(* IEC 61131-3 sources: helmsman/crates/helmsman-node/bench, 7 files *)

(* ---- analog_scale.st ---- *)
(* Raw analog count to engineering units, held to the range. bad is set when
   the raw value is outside raw_min..raw_max by more than the margin: a broken
   wire on a 4-20 mA loop, or a transmitter that has failed. *)
FUNCTION_BLOCK analog_scale
VAR_INPUT
  raw : REAL;
  raw_min : REAL := 0.0;
  raw_max : REAL := 32767.0;
  eng_min : REAL := 0.0;
  eng_max : REAL := 100.0;
  margin : REAL := 0.05;
END_VAR
VAR_OUTPUT
  value : REAL;
  bad : BOOL;
END_VAR
VAR
  span : REAL;
END_VAR
span := raw_max - raw_min;
bad := span <= 0.0 OR raw < raw_min - span * margin OR raw > raw_max + span * margin;
IF span > 0.0 THEN
  value := LIMIT(eng_min, eng_min + (raw - raw_min) / span * (eng_max - eng_min), eng_max);
END_IF;
END_FUNCTION_BLOCK

(* ---- batch_mixer.st ---- *)
(* Batch mixing tank: fill, heat while agitating, hold, drain, repeat.

   plant_model.st stands in for the tank so this runs with nothing wired. To
   wire real I/O: delete plant_model.st, delete the plant lines in the PROGRAM
   (each one says PLANT), and point io.map at your remote I/O module.

   A heater and agitator need a hardwired over-temperature cut-out and E-stop
   circuit. Those belong in hardware; nothing here is a safety function. *)

FUNCTION_BLOCK mixer_tank
VAR_INPUT
  run : BOOL;
  ack : BOOL;
  level_m : REAL;
  temp_c : REAL;
  inlet_open_sw : BOOL;
  inlet_closed_sw : BOOL;
  outlet_open_sw : BOOL;
  outlet_closed_sw : BOOL;
  agitator_fb : BOOL;
  agitator_overload : BOOL;
  overtemp_sw : BOOL;
END_VAR
VAR_OUTPUT
  inlet_coil : BOOL;
  outlet_coil : BOOL;
  agitator_contactor : BOOL;
  heater : BOOL;
  step : INT;
  batches : INT;
  tripped : BOOL;
  alarm_new : BOOL;
END_VAR
VAR CONSTANT
  fill_to_m : REAL := 2.0;        (* batch level *)
  empty_at_m : REAL := 0.05;      (* drained *)
  heater_min_m : REAL := 0.5;     (* element covered *)
  heat_to_c : REAL := 60.0;       (* batch temperature *)
  over_c : REAL := 80.0;          (* high temperature alarm *)
  hold_time : TIME := T#10s;      (* mix at temperature *)
  fill_max : TIME := T#60s;
  heat_max : TIME := T#120s;
  drain_max : TIME := T#60s;
END_VAR
VAR
  seq : step_sequencer;
  inlet : solenoid_valve;
  outlet : solenoid_valve;
  agitator : motor_starter;
  high_temp : latched_alarm;
  step_late : latched_alarm;
  equipment : latched_alarm;
  hold : TON;
  step_done : BOOL;
  step_max : TIME;
  want_inlet : BOOL;
  want_outlet : BOOL;
  want_agitator : BOOL;
  want_heat : BOOL;
END_VAR

high_temp(condition := overtemp_sw OR temp_c >= over_c, ack := ack, on_delay := T#0s);
step_late(condition := seq.timed_out, ack := ack, on_delay := T#0s);
equipment(condition := inlet.fault OR outlet.fault OR agitator.fault, ack := ack, on_delay := T#0s);
tripped := high_temp.showing OR step_late.showing OR equipment.showing;
alarm_new := high_temp.unacked OR step_late.unacked OR equipment.unacked;

seq(start := run AND NOT tripped, advance := step_done, abort := NOT run OR tripped,
    last_step := 4, step_limit := step_max);
step := seq.step;

want_inlet := FALSE;
want_outlet := FALSE;
want_agitator := FALSE;
want_heat := FALSE;
step_done := FALSE;
step_max := T#0s;
CASE step OF
  1: (* fill *)
    want_inlet := level_m < fill_to_m;
    step_done := level_m >= fill_to_m AND inlet.is_closed;
    step_max := fill_max;
  2: (* heat, agitating *)
    want_agitator := TRUE;
    want_heat := agitator.running;
    step_done := temp_c >= heat_to_c;
    step_max := heat_max;
  3: (* hold at temperature *)
    want_agitator := TRUE;
    want_heat := agitator.running AND temp_c < heat_to_c;
    step_done := hold.Q;
  4: (* drain *)
    want_outlet := level_m > empty_at_m;
    step_done := level_m <= empty_at_m AND outlet.is_closed;
    step_max := drain_max;
END_CASE;
hold(IN := step = 3, PT := hold_time);
IF seq.done AND batches < 32767 THEN
  batches := batches + 1;
END_IF;

inlet(open := want_inlet, at_open := inlet_open_sw, at_closed := inlet_closed_sw, reset := ack);
outlet(open := want_outlet, at_open := outlet_open_sw, at_closed := outlet_closed_sw, reset := ack);
agitator(run := want_agitator, feedback := agitator_fb, overload := agitator_overload, reset := ack);
inlet_coil := inlet.coil;
outlet_coil := outlet.coil;
agitator_contactor := agitator.contactor;
(* The heater never runs uncovered, without the agitator, or on an alarm. *)
heater := want_heat AND level_m >= heater_min_m AND NOT tripped;
END_FUNCTION_BLOCK

PROGRAM mixer
VAR_INPUT
  start_pb : BOOL;
  stop_pb : BOOL;
  ack_pb : BOOL;
  inlet_open_in : BOOL;
  inlet_closed_in : BOOL;
  outlet_open_in : BOOL;
  outlet_closed_in : BOOL;
  agitator_fb_in : BOOL;
  agitator_overload_in : BOOL;
  overtemp_in : BOOL;
  sim_inlet_stuck : BOOL;  (* PLANT: the inlet valve never opens *)
END_VAR
VAR_OUTPUT
  inlet_valve : BOOL;
  outlet_valve : BOOL;
  agitator : BOOL;
  heater : BOOL;
  lamp_green : BOOL;
  lamp_red : BOOL;
  step : INT;
  batches : INT;
  level_m : REAL;
  temp_c : REAL;
END_VAR
VAR
  plant : plant_model;  (* PLANT *)
  level_tx : analog_scale;
  temp_tx : analog_scale;
  tank : mixer_tank;
  light : stack_light;
  run : BOOL;
  level_raw : REAL;
  temp_raw : REAL;
  inlet_open : BOOL;
  inlet_closed : BOOL;
  outlet_open : BOOL;
  outlet_closed : BOOL;
  agitator_fb : BOOL;
END_VAR

plant(inlet := inlet_valve, outlet := outlet_valve, agitator := agitator, heater := heater,
      inlet_stuck := sim_inlet_stuck);  (* PLANT *)
level_raw := plant.level_raw;  (* PLANT: read your analog input here *)
temp_raw := plant.temp_raw;    (* PLANT: read your analog input here *)
inlet_open := inlet_open_in OR plant.inlet_open;  (* PLANT: keep the _in input *)
inlet_closed := inlet_closed_in OR plant.inlet_closed;  (* PLANT: keep the _in input *)
outlet_open := outlet_open_in OR plant.outlet_open;  (* PLANT: keep the _in input *)
outlet_closed := outlet_closed_in OR plant.outlet_closed;  (* PLANT: keep the _in input *)
agitator_fb := agitator_fb_in OR plant.agitator_fb;  (* PLANT: keep the _in input *)
run := (run OR start_pb) AND NOT stop_pb AND NOT tank.tripped;

level_tx(raw := level_raw, eng_min := 0.0, eng_max := 3.0);
temp_tx(raw := temp_raw, eng_min := 0.0, eng_max := 120.0);
tank(run := run, ack := ack_pb, level_m := level_tx.value, temp_c := temp_tx.value,
     inlet_open_sw := inlet_open, inlet_closed_sw := inlet_closed,
     outlet_open_sw := outlet_open, outlet_closed_sw := outlet_closed,
     agitator_fb := agitator_fb, agitator_overload := agitator_overload_in,
     overtemp_sw := overtemp_in);
light(running := run, alarm_new := tank.alarm_new, alarm_showing := tank.tripped);

inlet_valve := tank.inlet_coil;
outlet_valve := tank.outlet_coil;
agitator := tank.agitator_contactor;
heater := tank.heater;
lamp_green := light.green;
lamp_red := light.red;
step := tank.step;
batches := tank.batches;
level_m := level_tx.value;
temp_c := temp_tx.value;
END_PROGRAM

(* ---- latched_alarm.st ---- *)
(* One alarm: on after on_delay, stays showing until the condition has gone
   and someone has acknowledged it. *)
FUNCTION_BLOCK latched_alarm
VAR_INPUT
  condition : BOOL;
  ack : BOOL;
  on_delay : TIME;
END_VAR
VAR_OUTPUT
  active : BOOL;
  unacked : BOOL;
  showing : BOOL;
END_VAR
VAR
  delay : TON;
  rise : R_TRIG;
END_VAR
delay(IN := condition, PT := on_delay);
active := delay.Q;
rise(CLK := active);
IF rise.Q THEN
  unacked := TRUE;
ELSIF ack THEN
  unacked := FALSE;
END_IF;
showing := active OR unacked;
END_FUNCTION_BLOCK

(* ---- motor_starter.st ---- *)
(* Motor starter with contactor feedback and a latched fault.
   feedback is the contactor's auxiliary contact, overload the thermal relay.
   fault_code: 0 none, 1 overload, 2 no feedback after a start or feedback
   lost while running, 3 feedback with no command (contactor stuck on).
   A fault drops the contactor and holds until reset. An emergency stop
   belongs in a hardwired safety circuit, not in this block. *)
FUNCTION_BLOCK motor_starter
VAR_INPUT
  run : BOOL;
  feedback : BOOL;
  overload : BOOL;
  reset : BOOL;
  feedback_time : TIME := T#2s;
END_VAR
VAR_OUTPUT
  contactor : BOOL;
  running : BOOL;
  fault : BOOL;
  fault_code : INT;
END_VAR
VAR
  no_feedback : TON;
  stuck_on : TON;
END_VAR
no_feedback(IN := contactor AND NOT feedback, PT := feedback_time);
stuck_on(IN := NOT contactor AND feedback, PT := feedback_time);
IF overload THEN
  fault_code := 1;
ELSIF no_feedback.Q THEN
  fault_code := 2;
ELSIF stuck_on.Q THEN
  fault_code := 3;
ELSIF reset THEN
  fault_code := 0;
END_IF;
fault := fault_code <> 0;
contactor := run AND NOT fault;
running := contactor AND feedback;
END_FUNCTION_BLOCK

(* ---- solenoid_valve.st ---- *)
(* Single-solenoid valve or cylinder with an end switch each way.
   coil follows the command. fault latches when the switch for the commanded
   position has not made within travel_time, and clears on reset once the
   valve has arrived. Both switches on at once counts as not arrived. *)
FUNCTION_BLOCK solenoid_valve
VAR_INPUT
  open : BOOL;
  at_open : BOOL;
  at_closed : BOOL;
  reset : BOOL;
  travel_time : TIME := T#3s;
END_VAR
VAR_OUTPUT
  coil : BOOL;
  is_open : BOOL;
  is_closed : BOOL;
  fault : BOOL;
END_VAR
VAR
  late : TON;
END_VAR
coil := open;
is_open := at_open AND NOT at_closed;
is_closed := at_closed AND NOT at_open;
late(IN := (open AND NOT is_open) OR (NOT open AND NOT is_closed), PT := travel_time);
IF late.Q THEN
  fault := TRUE;
ELSIF reset THEN
  fault := FALSE;
END_IF;
END_FUNCTION_BLOCK

(* ---- stack_light.st ---- *)
(* Green while running. Red flashes for an alarm nobody has acknowledged and
   is steady for one that is acknowledged but still there. *)
FUNCTION_BLOCK stack_light
VAR_INPUT
  running : BOOL;
  alarm_new : BOOL;
  alarm_showing : BOOL;
END_VAR
VAR_OUTPUT
  green : BOOL;
  red : BOOL;
END_VAR
VAR
  flash : BLINK_PATTERN;
  pattern : INT;
END_VAR
IF alarm_new THEN
  pattern := 2;
ELSIF alarm_showing THEN
  pattern := 1;
ELSE
  pattern := 0;
END_IF;
flash(EN := TRUE, MODE := pattern, PERIOD := T#1s);
green := running;
red := flash.Q;
END_FUNCTION_BLOCK

(* ---- step_sequencer.st ---- *)
(* A numbered sequence. Step 0 is idle; start moves to step 1. Each step sets
   advance when it is finished, and the last step goes back to idle with done
   TRUE for one scan. step_limit is how long the current step may take (T#0s:
   no limit); past it, timed_out is set and the step holds until abort. abort
   returns to idle at once. Write the steps in a CASE on the step output. *)
FUNCTION_BLOCK step_sequencer
VAR_INPUT
  start : BOOL;
  advance : BOOL;
  abort : BOOL;
  last_step : INT;
  step_limit : TIME;
END_VAR
VAR_OUTPUT
  step : INT;
  step_time : TIME;
  timed_out : BOOL;
  done : BOOL;
END_VAR
VAR
  watch : TON;
  entered : BOOL;
END_VAR
done := FALSE;
entered := FALSE;
IF abort THEN
  step := 0;
  timed_out := FALSE;
  entered := TRUE;
ELSIF step = 0 THEN
  IF start THEN
    step := 1;
    entered := TRUE;
  END_IF;
ELSIF advance AND NOT timed_out THEN
  entered := TRUE;
  IF step >= last_step THEN
    step := 0;
    done := TRUE;
  ELSE
    step := step + 1;
  END_IF;
END_IF;
watch(IN := step > 0 AND NOT entered, PT := step_limit);
step_time := watch.ET;
IF step > 0 AND step_limit > T#0s AND watch.Q THEN
  timed_out := TRUE;
END_IF;
END_FUNCTION_BLOCK
